{attribute 'strict'}
{attribute 'qualified_only'}
TYPE E_ConveyorState : (Stopped := 0, Starting := 1, Running := 2, Fault := 3);
END_TYPE

(* stored: Version 1.1.0.1, ProductVersion 3.1 *)
